PROGRAM SerialBackground
VAR
	fbDomeSerial : FB_SerialBackground;
	fbPendantSerial : FB_SerialBackground;
END_VAR

fbDomeSerial(RxBuffer:=RxBufferDome, TxBuffer:=TxBufferDome);

fbPendantSerial(RxBuffer:=RxBufferPendant, TxBuffer:=TxBufferPendant);

END_PROGRAM

(* stored: Version 1.1.0.1, ProductVersion 3.1.4024.15
   POU SerialBackground: Id {9a20473f-0d3f-4584-b429-33e10587a848}, SpecialFunc None *)
